Fanuc KAREL source: kb00024.KL

PROGRAM KB00024
%NOLOCKGROUP
VAR
P1 : FILE
BEGIN
CLR_IO_STAT(P1)
END KB00024
